RESOURCE RES0 : EMB_RES_ECO
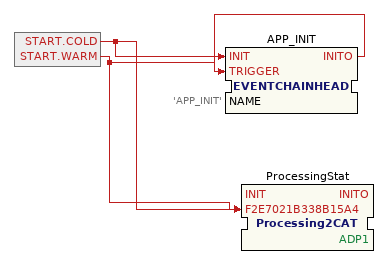
  FBS
    APP_INIT : EVENTCHAINHEAD(NAME := 'APP_INIT');
    ProcessingStat : Processing2CAT;
  END_FBS
  EVENT_CONNECTIONS
    START.COLD TO APP_INIT.INIT;
    START.WARM TO APP_INIT.INIT;
    APP_INIT.INITO TO APP_INIT.TRIGGER;
    START.COLD TO ProcessingStat.F2E7021B338B15A4;
    START.WARM TO ProcessingStat.F2E7021B338B15A4;
  END_CONNECTIONS
END_RESOURCE
